Fanuc KAREL source: KT00797.KL

PROGRAM KT00797
%NOLOCKGROUP
VAR
  I1: INTEGER
  I2: INTEGER
  OUT: REAL
BEGIN
  I1 = 2
  I2 = 3
  I1 = 2
  I2 = 3
  OUT = EXP(I1)
END KT00797
